Staubli VAL3: utContainer.pjx

--- utContainer.pjx ---
Parameters version=s8.8.3Cs9_BS1660 stackSize=5000 millimeterUnit=true
Program file=start.pgx
Program file=stop.pgx
Data file=utContainer.dtx
Type name=utAppearance path=./utAppearance/utAppearance.pjx
Type name=utCommon path=./utCommon/utCommon.pjx

--- utContainer.dtx ---
public utAppearance Appearance
  [0]
    bool bVisibility
public utCommon Common
  [0]
    string sSource
    string sID
    string sPage

--- start.pgx ---
program start()
begin
end

--- stop.pgx ---
program stop()
begin
end
